Fanuc KAREL source: KT00131.KL

PROGRAM KT00131
%NOLOCKGROUP
VAR
  I1: INTEGER
  R2: REAL
  OUT: INTEGER
BEGIN
  I1 = 2
    R2 = 3.0
  OUT = I1 DIV R2
END KT00131
